{attribute 'qualified_only'}
{attribute 'strict'}
{attribute 'to_string'}
TYPE E_LogRecordProcessorFailureReason :
(
	NA := 0,  // No failure occurred.
	RECORD_CLONE_FAILURE,  // The emitted record could not be cloned for retention.
	QUEUE_PUSH_FAILURE,  // The retained record could not be transferred into the queue.
	EXPORT_FAILURE  // The exporter did not accept the prepared batch.
) UDINT;
END_TYPE

(* stored: Version 1.1.0.1
   EnumerationTextList E_LogRecordProcessorFailureReason: Id {d584c2c7-6b3c-46ad-8152-e53006c991ce} *)
